// TIA Portal V19 export
// export: Created 2026-10-15T10:10:35.3496691Z, ExportSetting WithDefaults, DisplayName Totally Integrated Automation Portal, DisplayVersion V19, DisplayName TIA Portal Openness, DisplayVersion V19, DisplayName TIA Portal Version Control Interface, DisplayVersion V19, DisplayName STEP 7 Professional, DisplayVersion V19, DisplayName STEP 7 Safety, DisplayVersion V19, DisplayName WinCC Basic/Comfort/Advanced, DisplayVersion V19, DisplayName WinCC Unified, DisplayVersion V19
FUNCTION "ROLL_PB3" : Void   // FC15, SCL
{ S7_Optimized_Access := 'TRUE' }
VERSION : 0.1
// stored: AutoNumber true, IsIECCheckEnabled false, SetENOAutomatically false, UDAEnableTagReadback false
   VAR_TEMP
      r : Bool;
      a1 : Word;
      a2 : Word;
      activeDataBlock : Int;
      comparisonResults : Array[0..15] of Bool;
   END_VAR
BEGIN

   #r := FALSE;
   #a1 := W#16#0000;
   #a2 := W#16#0000;
   #activeDataBlock := 0;
   // PB3, STEP 5 network 1
   #a2 := #a1;
   #a1 := "ROLL_GetM"(FirstByte := 239, Width := 8);
   #a2 := #a1;
   #a1 := W#16#0001;
   #comparisonResults[0] := (WORD_TO_INT(#a2) = WORD_TO_INT(#a1));
   #r := #comparisonResults[0];
   "ROLL_State".M[20, 1] := #r;
   // PB3, STEP 5 network 2
   #a2 := #a1;
   #a1 := "ROLL_GetM"(FirstByte := 239, Width := 8);
   #a2 := #a1;
   #a1 := W#16#0002;
   #comparisonResults[1] := (WORD_TO_INT(#a2) = WORD_TO_INT(#a1));
   #r := #comparisonResults[1];
   "ROLL_State".M[20, 2] := #r;
   // PB3, STEP 5 network 3
   #a2 := #a1;
   #a1 := "ROLL_GetM"(FirstByte := 239, Width := 8);
   #a2 := #a1;
   #a1 := W#16#0003;
   #comparisonResults[2] := (WORD_TO_INT(#a2) = WORD_TO_INT(#a1));
   #r := #comparisonResults[2];
   "ROLL_State".M[20, 3] := #r;
   // PB3, STEP 5 network 4
   #a2 := #a1;
   #a1 := "ROLL_GetM"(FirstByte := 239, Width := 8);
   #a2 := #a1;
   #a1 := W#16#0004;
   #comparisonResults[3] := (WORD_TO_INT(#a2) = WORD_TO_INT(#a1));
   #r := #comparisonResults[3];
   "ROLL_State".M[20, 4] := #r;
   // PB3, STEP 5 network 5
   #a2 := #a1;
   #a1 := "ROLL_GetM"(FirstByte := 239, Width := 8);
   #a2 := #a1;
   #a1 := W#16#0005;
   #comparisonResults[4] := (WORD_TO_INT(#a2) = WORD_TO_INT(#a1));
   #r := #comparisonResults[4];
   "ROLL_State".M[20, 5] := #r;
   // PB3, STEP 5 network 6
   #a2 := #a1;
   #a1 := "ROLL_GetM"(FirstByte := 239, Width := 8);
   #a2 := #a1;
   #a1 := W#16#0007;
   #comparisonResults[5] := (WORD_TO_INT(#a2) = WORD_TO_INT(#a1));
   #r := #comparisonResults[5];
   "ROLL_State".M[20, 7] := #r;
   // PB3, STEP 5 network 7
   #a2 := #a1;
   #a1 := "ROLL_GetM"(FirstByte := 239, Width := 8);
   #a2 := #a1;
   #a1 := W#16#000A;
   #comparisonResults[6] := (WORD_TO_INT(#a2) = WORD_TO_INT(#a1));
   #r := #comparisonResults[6];
   "ROLL_State".M[22, 0] := #r;
   // PB3, STEP 5 network 8
   #a2 := #a1;
   #a1 := "ROLL_GetM"(FirstByte := 239, Width := 8);
   #a2 := #a1;
   #a1 := W#16#000B;
   #comparisonResults[7] := (WORD_TO_INT(#a2) = WORD_TO_INT(#a1));
   #r := #comparisonResults[7];
   "ROLL_State".M[22, 1] := #r;
   // PB3, STEP 5 network 9
   #a2 := #a1;
   #a1 := "ROLL_GetM"(FirstByte := 239, Width := 8);
   #a2 := #a1;
   #a1 := W#16#000C;
   #comparisonResults[8] := (WORD_TO_INT(#a2) = WORD_TO_INT(#a1));
   #r := #comparisonResults[8];
   "ROLL_State".M[22, 2] := #r;
   // PB3, STEP 5 network 10
   #a2 := #a1;
   #a1 := "ROLL_GetM"(FirstByte := 239, Width := 8);
   #a2 := #a1;
   #a1 := W#16#000D;
   #comparisonResults[9] := (WORD_TO_INT(#a2) = WORD_TO_INT(#a1));
   #r := #comparisonResults[9];
   "ROLL_State".M[22, 3] := #r;
   // PB3, STEP 5 network 11
   #a2 := #a1;
   #a1 := "ROLL_GetM"(FirstByte := 239, Width := 8);
   #a2 := #a1;
   #a1 := W#16#000E;
   #comparisonResults[10] := (WORD_TO_INT(#a2) = WORD_TO_INT(#a1));
   #r := #comparisonResults[10];
   "ROLL_State".M[22, 4] := #r;
   // PB3, STEP 5 network 12
   #a2 := #a1;
   #a1 := "ROLL_GetM"(FirstByte := 239, Width := 8);
   #a2 := #a1;
   #a1 := W#16#000F;
   #comparisonResults[11] := (WORD_TO_INT(#a2) = WORD_TO_INT(#a1));
   #r := #comparisonResults[11];
   "ROLL_State".M[22, 5] := #r;
   // PB3, STEP 5 network 13
   #a2 := #a1;
   #a1 := "ROLL_GetM"(FirstByte := 239, Width := 8);
   #a2 := #a1;
   #a1 := W#16#0014;
   #comparisonResults[12] := (WORD_TO_INT(#a2) = WORD_TO_INT(#a1));
   #r := #comparisonResults[12];
   "ROLL_State".M[23, 0] := #r;
   // PB3, STEP 5 network 14
   #a2 := #a1;
   #a1 := "ROLL_GetM"(FirstByte := 239, Width := 8);
   #a2 := #a1;
   #a1 := W#16#0015;
   #comparisonResults[13] := (WORD_TO_INT(#a2) = WORD_TO_INT(#a1));
   #r := #comparisonResults[13];
   "ROLL_State".M[23, 1] := #r;
   // PB3, STEP 5 network 15
   #a2 := #a1;
   #a1 := "ROLL_GetM"(FirstByte := 239, Width := 8);
   #a2 := #a1;
   #a1 := W#16#0016;
   #comparisonResults[14] := (WORD_TO_INT(#a2) = WORD_TO_INT(#a1));
   #r := #comparisonResults[14];
   "ROLL_State".M[23, 2] := #r;
   // PB3, STEP 5 network 16
   #a2 := #a1;
   #a1 := "ROLL_GetM"(FirstByte := 239, Width := 8);
   #a2 := #a1;
   #a1 := W#16#0017;
   #comparisonResults[15] := (WORD_TO_INT(#a2) = WORD_TO_INT(#a1));
   #r := #comparisonResults[15];
   "ROLL_State".M[23, 3] := #r;
   // PB3, STEP 5 network 17
   RETURN;
END_FUNCTION
